// Model of the TwinSAFE FB RS (reset dominant latch).
// The Safety Editor refuses an RS with Set or Reset unconnected: the model then reports Error with
// diagnostic bit 15 instead of running (see T_SafeFunctionBlockBase).
{attribute 'reflection'}
FUNCTION_BLOCK T_SafeRs EXTENDS T_SafeFunctionBlockBase
VAR_INPUT
    Set : BOOL;
    Reset : BOOL;
    Parameters : ST_SafeLatchParameters;
END_VAR
VAR_OUTPUT
    RsOut : BOOL;
END_VAR
VAR
    {attribute 'is_connected' := 'Set'}
    _setConnected : BOOL;
    {attribute 'is_connected' := 'Reset'}
    _resetConnected : BOOL;
    _state : E_SafeLatchState := E_SafeLatchState.Stop;
END_VAR

SUPER^();

// Set and Reset must both be connected (Safety Editor: "Inport Set of RS must be connected").
METHOD PROTECTED ConfigurationOk : BOOL
IF NOT _setConnected THEN
    _configurationFault := 'T_SafeRs: Inport Set of RS must be connected';
    RETURN;
ELSIF NOT _resetConnected THEN
    _configurationFault := 'T_SafeRs: Inport Reset of RS must be connected';
    RETURN;
END_IF

ConfigurationOk := TRUE;
END_METHOD

METHOD PROTECTED Process
VAR
    setActive : BOOL;
    resetActive : BOOL;
END_VAR
setActive   := F_SafeInputValue(_setConnected, Parameters.SetMakeContact, Set);
resetActive := F_SafeInputValue(_resetConnected, Parameters.ResetMakeContact, Reset);

IF NOT _fbRun THEN
    _state := E_SafeLatchState.Stop;
ELSE
    IF _state = E_SafeLatchState.Stop THEN
        _state := E_SafeLatchState.Safe;
    END_IF

    IF resetActive THEN
        _state := E_SafeLatchState.Safe;
    ELSIF setActive THEN
        _state := E_SafeLatchState.Set;
    END_IF
END_IF

RsOut := (_state = E_SafeLatchState.Set);
Error := FALSE;
Diag  := 0;
State := TO_BYTE(_state);
END_METHOD

END_FUNCTION_BLOCK

(* stored: Version 1.1.0.1
   POU T_SafeRs: Id {e620cd2a-846a-5dd3-8008-ec245bc27373}, SpecialFunc None
   Method ConfigurationOk: Id {d0a116af-3fb8-47bb-be2e-5d59e9963190}
   Method Process: Id {84936541-d311-5217-9cf7-620653b0d636} *)
